// System API/DSM/API/bds_dsm_getDFES_DTC
///This function is used to get DTC values and total number of errors present in DFES entry.
///
///=======
/// Remarks:
///=======
///    + The |GVL_dsm| is given for usage of defines.
///
///----------
/// FFI:
///----------
///This API can be used in trusted partitions only. See Freedom from Interference (FFI) concept for more details.
///
///-----
/// NOTICE:
///-----
///    + On a maximum, 32 different DFES entries are possible. 
///    + Status Mask will take time (max. 10ms) to update in global mask so return status has to be monitored.
///	
///==================================================================		  			===================================================================================================
///Return value    								  									Description
///==================================================================		  			===================================================================================================
///16#0000: BDS_DSM_NO_ERROR_DU16														Update of DTC values and total number of errors present is successful .
///16#0004: BDS_DSM_INVALID_PTR_DU16													Invalid Pointer.
///16#0005: BDS_DSM_MASK_ERROR_DU16													Invalid Mask.
///16#0007: BDS_DSM_INVALID_MAX_ERROR_DU16 											Invalid Max Error.
///16#000B: BDS_DSM_NO_DTC_AVAILABLE_DU16 												Invalid DTC value.
///
///==================================================================		   			===================================================================================================
///
///
///=======
///Code Example:
///=======
///============================================================================
///
///PROGRAM BDS_DSM_getDFES_DTC_TEST
///
///VAR
///
///	mask_s : UINT := BDS_DSM_SET_ACTIVE_ERROR_MASK_DU16;
///
///	startFromBegin_l: BOOL := TRUE;
///
///	maxNum_u16:UINT := 32;
///
///	error_count_u16: UINT;
///
///	dtc_pu16: ARRAY [1..32] OF UINT;
///
///	status_u16: UINT;
///
///END_VAR
///
///dfc_s.id := dfc_ts.DFCid;
///
///(*Get DFES entries*)
///
///status_u16 := bds_dsm_getDFES(mask_s, TRUE, maxNum_u16, ADR(error_count_u16), ADR(dtc_pu16));
///
///if status_u16 = BDS_DSM_NO_ERROR_DU16 THEN
///
///	(*Numbers of Errors have been read successfully*)
///
///END_IF
///
///============================================================================
///
{attribute 'external_name' := 'cmp_rts_bds_dsm_getDFES_DTC'}
FUNCTION bds_dsm_getDFES_DTC : UINT
VAR_INPUT
	///The kind of error status can be specified in detail by means of this mask.
	///
	///Possible values:
	///    + BDS_DSM_SET_ACTIVE_ERROR_MASK_DU16 ( 16#18 ) - Fault is active.
	///    + BDS_DSM_SET_TESTED_ONCE_MASK_DU16 ( 16#08 ) - DFC was tested at least once since start or reset.
	///    + BDS_DSM_SET_TESTED_OK_MASK_DU16 ( 16#20 ) - DFC was at least once ok tested since start or reset.  
	///    + BDS_DSM_SET_FAILED_SINCE_CLEAR_MASK_DU16 ( 16#80 ) - Fault occured at least once since error was deleted from memory.
	mask_s: UINT;
	///
	///    + TRUE: Query is started from the beginning of DFES.
	///    + FALSE: Query is continued with the next index where the last query was finished.
	startFromBegin_l: BOOL;
	///Maximal number of errors/DTCs is returned. The BSW will return at max. 32 values (the max. size of DFES).
	maxNum_u16: UINT;
	///Pointer to a variable where the total number of errors is returned.
	num_pu16: POINTER TO UINT;
	///Pointer variable used to store DTC values.
	dtc_pu16: POINTER TO UINT;
END_VAR

END_FUNCTION

// System API/DSM/API/bds_dsm_getDTC_DFC
///This function returns the DTC of a specified DFC.
///
///=======
/// Remarks:
///=======
///    + The |GVL_dsm| is given for usage of defines.
///	
///----------
/// FFI:
///----------
///This API can be used in trusted partitions only. See Freedom from Interference (FFI) concept for more details.
///
///==================================================================		  			===================================================================================================
///Return value    								  									Description
///==================================================================		  			===================================================================================================
///16#0000: BDS_DSM_NO_ERROR_DU16														Update of DTC of DFC is Successful .
///16#0001: BDS_DSM_DFC_ERROR_DU16														Invalid DFC.
///16#0004: BDS_DSM_INVALID_PTR_DU16													Invalid pointer.
///
///==================================================================		   			===================================================================================================
///
///
///=======
///Code Example:
///=======
///============================================================================
///
///PROGRAM bds_dsm_getDTC_DFC_TEST
///
///VAR
///
///	dfc_s: bds_dsm_dfc_ts;	
///
///	dfc_ts : DFC_bds_NoDebFault1;
///
///	dtc_error_u16 : UINT;
///
///	status_u16: UINT;
///
///END_VAR
///
///dfc_s.id := dfc_ts.DFCid;
///
///(*Read the DTC of DFC*)
///
///dfc_s.id := dfc_ts.DFCid;
///
///status_u16 := bds_dsm_getDTC_DFC(dfc_s,ADR(dtc_error_u16));
///
///if status_u16 = BDS_DSM_NO_ERROR_DU16 THEN
///
///	(*DTC of DFC was read successful*)
///
///END_IF
///
///============================================================================
///
{attribute 'external_name' := 'cmp_rts_bds_dsm_getDTC_DFC'}
FUNCTION bds_dsm_getDTC_DFC : UINT
VAR_INPUT
	///DFC name (identifier) : It is configured using easyConfig tool.
	dfc_s: bds_dsm_dfc_ts;
	///Pointer to a variable where the DTC is returned.
	dtc_pu16: POINTER TO UINT;
END_VAR

END_FUNCTION

// System API/DSM/API/bds_dsm_getDTC_DFCJ1939
///This function is used to read the J1939 specific DTC data (SPN, FMI, Lamp states) for a given DFC.
///
///=======
/// Remarks:
///=======
///    + The |GVL_dsm| is given for usage of defines.
///	+ Suspect Parameter Number (SPN), Failure Mode Identifier (FMI) and Lamp States can be configured in easyConfig.
///	
///----------
/// FFI:
///----------
///This API can be used in trusted partitions only. See Freedom from Interference (FFI) concept for more details.
///
///==================================================================		  			===================================================================================================
///Return value    								  									Description
///==================================================================		  			===================================================================================================
///16#0000: BDS_DSM_NO_ERROR_DU16														Read data is successful.
///16#0001: BDS_DSM_DFC_ERROR_DU16														Wrong DFC.
///16#0004: BDS_DSM_INVALID_PTR_DU16													Invalid Pointer.
///
///==================================================================		   			===================================================================================================
///
///
///=======
///Code Example:
///=======
///============================================================================
///
///PROGRAM bds_dsm_getDTC_DFCJ1939_TEST
///
///VAR
///
///	dfc_s: bds_dsm_dfc_ts;	
///
///	dfc_ts : DFC_bds_NoDebFault1;
///
///	dtcJ1939_s : bds_dsm_dtcj1939_ts;
///
///	status_u16: UINT;
///
///END_VAR
///
///dfc_s.id := dfc_ts.DFCid;
///
///(*Read the DTC of DFC*)
///
///dfc_s.id := dfc_ts.DFCid;
///
///status_u16 := bds_dsm_getDTC_DFCJ1939(dfc_s, ADR(dtcJ1939_s));
///
///if status_u16 = BDS_DSM_NO_ERROR_DU16 THEN
///
///	(*J1939 specific DTC data is read successfull*)
///
///END_IF
///
///============================================================================
///
{attribute 'external_name' := 'cmp_rts_bds_dsm_getDTC_DFCJ1939'}
FUNCTION bds_dsm_getDTC_DFCJ1939 : UINT
VAR_INPUT
	///DFC name (identifier) : It is configured using easyConfig tool.
	dfc_s: bds_dsm_dfc_ts;
	///pointer to a variable where the DTC data is returned.
	dtcJ1939_ps: POINTER TO bds_dsm_dtcj1939_ts;
END_VAR

END_FUNCTION

// System API/DSM/API/bds_dsm_getDTC_J1939
///This function is used to read the J1939 specific DTC data (SPN, FMI, Lamp states) for a given DTC.
///
///=======
/// Remarks:
///=======
///    + The |GVL_dsm| is given for usage of defines.
///	+ Suspect Parameter Number (SPN), Failure Mode Identifier (FMI) and Lamp States can be configured in easyConfig.
///	
///----------
/// FFI:
///----------
///This API can be used in trusted partitions only. See Freedom from Interference (FFI) concept for more details.
///
///----------
/// FFI:
///----------
///This API can be used in trusted partitions only. See Freedom from Interference (FFI) concept for more details.
///
///==================================================================		  			===================================================================================================
///Return value    								  									Description
///==================================================================		  			===================================================================================================
///16#0000: BDS_DSM_NO_ERROR_DU16														Update of J1939 specific data is successful .
///16#0004: BDS_DSM_INVALID_PTR_DU16													Invalid Pointer.
///16#000B: BDS_DSM_NO_DTC_AVAILABLE_DU16												Invalid DTC input.
///
///==================================================================		   			===================================================================================================
///
///
///=======
///Code Example:
///=======
///============================================================================
///
///PROGRAM DSM
///
///VAR
///
///	dfc_s: bds_dsm_dfc_ts;
///
///	dfc_ts : DFC_bds_NoDebFault1;
///
///	dtcJ1939_s: bds_dsm_dtcj1939_ts;
///
///	dtc_u16:UINT := 32772;
///
///	status_u16: UINT;
///
///END_VAR
///
///dfc_s.id := dfc_ts.DFCid;
///
///(*Read the DTC of DFC*)
///
///dfc_s.id := dfc_ts.DFCid;
///
///status_u16 := bds_dsm_getDTC_J1939(dtc_u16, ADR(dtcJ1939_s));
///
///if status_u16 = BDS_DSM_NO_ERROR_DU16 THEN
///
///	(*J1939 specific DTC data is read successfull*)
///
///END_IF
///
///============================================================================
///
///
{attribute 'external_name' := 'cmp_rts_bds_dsm_getDTC_J1939'}
FUNCTION bds_dsm_getDTC_J1939 : UINT
VAR_INPUT
	///DTC value : It is configured using easyConfig tool.
	dtc_u16: UINT;
	///pointer to a variable where the DTC data is returned.
	dtcJ1939_ps: POINTER TO bds_dsm_dtcj1939_ts;
END_VAR

END_FUNCTION

// I/O API/IN legacy/API/bds_in_fi_buffered
///Provides the period array and pulse array of a frequency signal.
///
///=======
/// Remarks:
///=======
///   + In order to receive  the buffered frequency of a signal, it should be configured with easyConfig as a frequency signal. Once configured it is automatically enabled during the start up of the ECU.
///   + For information about the signal acquisition see Frequency acquisition.
///   + If application uses an invalid channel  as a parameter while calling the function, the values stored in the data structure will be 0 // replacement
///   + The following signal information is available: 
///	   + Pointer to the starting address of the Period array (Max size 20).
///	   + Pointer to the starting address of Pulse array (Max size 20).
///   + After the function is called  you get  20  samples of periods and pulses  that could be used within a loop.  
///
///
///----------
/// FFI:
///----------
///This API can be used in trusted partitions only. See Freedom from Interference (FFI) concept for more details.
///
///==================================================================		  			===================================================================================================
///Return value    								  									Description
///==================================================================		  			===================================================================================================
///0																					No error
///1																					Invalid parameter
///2																					Function call was erroneous
///
///==================================================================		   			===================================================================================================
{attribute 'external_name' := 'cmp_rts_bds_in_fi_buffered'}
FUNCTION bds_in_fi_buffered : USINT
VAR_INPUT
	///The signal name that is assigned to the respective pin configured as frequency input. see bds_in_fi_signal_te in bds_rts_ec.xml
	signal_e: UINT;
	///POINTER TO |bds_in_FrqBuffered_ts|
	data_ps: POINTER TO bds_in_FrqBuffered_ts;
END_VAR

END_FUNCTION

// System API/SYS/API/bds_sysPb_getVariant
///This function gets the currently selected post-build selectable variant.
///
///Refer to the page Post-build selectable for more information.
///
///=======
/// Remarks:
///=======
///    + The |GVL_sys| is given for usage of defines.
///    + This Api should be called once in application
///
///----------
/// FFI:
///----------
///This API can be used in trusted partitions.  For untrusted partitions use |bds_sysPb_getVariant_ffi|. See Freedom from Interference (FFI) concept for more details.
///
///==================================================================		  			===================================================================================================
///Return value    								  									Description
///==================================================================		  			===================================================================================================
///|bds_sysPb_retValGetVrnt_ts|															Currently configured variant.
///
///==================================================================		   			===================================================================================================
///
///=======
///Code Example:
///=======
///============================================================================
///
///PROGRAM IniProc
///
///VAR
///	getVaraint_s: bds_sysPb_retValGetVrnt_ts;
///END_VAR
///
///(*getVaraint_s contains the current selected variant*)
///
///getVaraint_s = bds_sysPb_getVariant();
///
///============================================================================
{attribute 'external_name' := 'cmp_rts_bds_sysPb_getVariant'}
FUNCTION bds_sysPb_getVariant : bds_sysPb_retValGetVrnt_ts

END_FUNCTION

// System API/SYS/FFI_API/bds_sysPb_getVariant_ffi
{attribute 'external_name' := 'cmp_rts_bds_sysPb_getVariant_ffi'}
FUNCTION bds_sysPb_getVariant_ffi : bds_sysPb_retValGetVrnt_ts

END_FUNCTION

// System API/SYS/API/bds_sysPb_cfgVariant
///This function is used to select desired variant in the ECU.
///
///Refer to the page Post-build selectable for more information.
///
///=======
/// Remarks:
///=======
///
///The |GVL_sys| is given for usage of defines.
///The selected variant will take effect only after one of the following actions,
///    + A soft reset via bds_sys_resetECU.
///    + Ignition OFF and ON.
///
///----------
/// FFI:
///----------
///This API can be used in trusted partitions only. See Freedom from Interference (FFI) concept for more details.
///
///----------
/// NOTICE:
///----------
///    + The selectable variants will be listed in bds_sysPb_vrnt_te.Import the bds_rts_ec.xml to use the enum.
///    + The configuration related to the particular variant has to be looked-up in easyConfig.
///    + As of now IN module is alone supported for Post-build selectable.
///
///==================================================================		  			===================================================================================================
///Return value    								  									Description
///==================================================================		  			===================================================================================================
///16#0																					No errors, API executed successfully.New variant is updated in RAM successfully.
///16#1																					Invalid variant input.
///16#2																					Variant is already selected
///==================================================================		   			===================================================================================================
///
///=======
///Code Example:
///=======
///============================================================================
///
///PROGRAM IniProc
///
///VAR
///	statusCfgVrnt_s: bds_sysPb_retValCfgVrnt_ts;
///	cfgPbVrnt_u8:usint:=0;
///
///END_VAR
///
///(*Configure a variant. eg bds_sysPb_vrnt03_E*)
///(*Call API once*)
///IF(0 = cfgPbVrnt_u8) THEN
///
///	statusCfgVrnt_s:=bds_sysPb_cfgVariant(bds_sysPb_vrnt_te.bds_sysPb_vrnt03_E);
///
///(*do ignition OFF & ON or do soft reset via bds_sys_resetECU.*)
///cfgPbVrnt_u8:=1;
///
///END_IF
///============================================================================
{attribute 'external_name' := 'cmp_rts_bds_sysPb_cfgVariant'}
FUNCTION bds_sysPb_cfgVariant : bds_sysPb_retValCfgVrnt_ts
VAR_INPUT
	vrntParam_e: USINT;
END_VAR

END_FUNCTION

// I/O API/SENT/API/bds_sent_getFastData
(*The bds_sent_getFastData API function provides the received SENT Fast Data of the selected input signal.

=======
 Remarks:
=======
    + Before accessing the Fast Data frame, check the function call status in the return data structure |bds_sent_rxFastData_ts|.
    + If the function call status is bds_sentCmn_ok_E, then the received Fast Data nibbles from array rxFastData_au8 in the return data structure |bds_sent_rxFastData_ts| can be used. Otherwise the data is set to zero.
    + The function call will return a negative response code if a false parameter is used (e.g., selected signal_e is not defined as SENT input signal or is not configured in Post-Build-Selectable variant).
	+ The positive or negative response codes (e.g., bds_sentCmn_ok_E, bds_sentCmn_notAvl_E and bds_sentCmn_errExt_E) provide in the return data structure |bds_sent_rxFastData_ts| a detailed SENT driver status information chSt_b in bit format.
	+ The number of received Fast Data Nibbles per frame can be configured in easyConfig with the value bds_sent_maxDataNibbles_du8.
	+ The value of the macro define bds_sent_maxDataNibbles_du8 depends on the selected SENT J2716 protocol version. The possible values that can be set in easyConfig are 6 or 8 data nibbles.
	+ The entire SENT channel-specific configuration is to be performed in easyConfig.
	+ Decoding of SENT data is not provided by the API function.

----------
 FFI:
----------
This API can be used in trusted partitions . For untrusted partitions use |bds_sent_getFastData_ffi|. See Freedom from Interference (FFI) concept for more details.
	
==================================================================		  			===================================================================================================
Return value    								  									Description
==================================================================		  			===================================================================================================
|bds_sent_rxFastData_ts|															The return data structure containing the latest received Fast Data sample and the state information.

==================================================================		   			===================================================================================================

=======
Code Example:
=======
============================================================================

PROGRAM appl_10ms_task
VAR

	bds_sent_rxFastData_s : bds_sent_rxFastData_ts;

	idx:USINT;

	appl_sent_rxFastData_au8: ARRAY[1..8] OF USINT;	
	
END_VAR

// Get the single Fast Data frame on selected SENT signal K59

 bds_sent_rxFastData_s = bds_sent_getFastData(bds_sent_signal_te.bds_sent_K59_E);
 
IF(bds_sentCmn_ok_E = bds_sent_rxFastData_s.status_e) THEN
 
    IF(1 = bds_sent_rxFastData_s.chSt_b.newFrmRxd_b1) THEN
   
      // Save the new received Fast Data frame.

      // Received data nibbles saved in low nibble of byte array element (high data nibble set to "0".

		FOR idx := 1 TO 8 BY 1 DO

			appl_sent_rxFastData_au8[idx] := bds_sent_rxFastData_s.rxFastData_au8[idx];

		END_FOR;

    END_IF
  
END_IF

============================================================================

*)
{attribute 'external_name' := 'cmp_rts_bds_sent_getFastData'}
FUNCTION bds_sent_getFastData : bds_sent_rxFastData_ts
VAR_INPUT
	(*The signal name that is assigned to the respective pin configured as SENT channel*)
	signal_e: USINT;
END_VAR

END_FUNCTION

// I/O API/SENT/FFI_API/bds_sent_getFastData_ffi
{attribute 'external_name' := 'cmp_rts_bds_sent_getFastData_ffi'}
FUNCTION bds_sent_getFastData_ffi : bds_sent_rxFastData_ts
VAR_INPUT
	(*The signal name that is assigned to the respective pin configured as SENT channel*)
	signal_e: USINT;
END_VAR

END_FUNCTION

// I/O API/SENT/API/bds_sent_getSlowData
(*The bds_sent_getSlowData API function provides the received SENT Slow Data of the selected input signal.

=======
 Remarks:
=======
    + Before accessing the Slow Data frame, check the function call status in the return data structure |bds_sent_rxSlowData_ts|.
    + If the function call status is bds_sentCmn_ok_E, then the received Slow Data messages from element rxSlowData_u32, msgId_u8 and cfgBit_u8 in the return data structure |bds_sent_rxSlowData_ts| can be used. Otherwise the data is set to zero.
	+ The function call will return a negative response code if a false parameter is used (e.g. selected signal_e is not defined as SENT input signal or is not configured in Post-Build-Selectable variant).
	+ The positive or negative response codes bds_sentCmn_ok_E, bds_sentCmn_notAvl_E and bds_sentCmn_errExt_E support in the return data structure |bds_sent_rxSlowData_ts| a detailed SENT driver status information chSt_b in bit format.
	+ The entire SENT channel-specific configuration is to be performed in easyConfig.
	+ Decoding of SENT data is not provided by the API function.

----------
 FFI:
----------
This API can be used in trusted partitions . For untrusted partitions use |bds_sent_getSlowData_ffi|. See Freedom from Interference (FFI) concept for more details.
	
==================================================================		  			===================================================================================================
Return value    								  									Description
==================================================================		  			===================================================================================================
|bds_sent_rxSlowData_ts|															The return data structure containing the latest received Slow Data sample and the state information

==================================================================		   			===================================================================================================

=======
Code Example:
=======
============================================================================

PROGRAM appl_10ms_task
VAR

	bds_sent_rxSlowData_s : bds_sent_rxSlowData_ts;

	rxSlowData_u32:UDINT;

	SlowData_msgId_u8: USINT;	
	
	SlowData_cfgBit_u8: USINT;
	
END_VAR

// Get the single Slow Data frame on selected SENT signal K59

  bds_sent_rxSlowData_s = bds_sent_getSlowData(bds_sent_signal_te.bds_sent_K59_E);
 
IF(bds_sentCmn_ok_E = bds_sent_rxSlowData_s.status_e) THEN
	
	//Get SENT status information if new Slow Data frame received
 
    IF(1 = bds_sent_rxSlowData_s.chSt_b.newSlowFrmRxd_b1) THEN
   
      // Save the new received Slow Data frame

		rxSlowData_u32 := bds_sent_rxSlowData_s.rxSlowData_u32;

		SlowData_msgId_u8 := bds_sent_rxSlowData_s.msgId_u8;
		
		SlowData_cfgBit_u8 := bds_sent_rxSlowData_s.cfgBit_u8;

	  ELSE

		//error handling for no new Slow Data frame received

    END_IF
  
END_IF

============================================================================

*)
{attribute 'external_name' := 'cmp_rts_bds_sent_getSlowData'}
FUNCTION bds_sent_getSlowData : bds_sent_rxSlowData_ts
VAR_INPUT
	(*The signal name that is assigned to the respective pin configured as SENT channel*)
	signal_e: USINT;
END_VAR

END_FUNCTION

// I/O API/SENT/FFI_API/bds_sent_getSlowData_ffi
{attribute 'external_name' := 'cmp_rts_bds_sent_getSlowData_ffi'}
FUNCTION bds_sent_getSlowData_ffi : bds_sent_rxSlowData_ts
VAR_INPUT
	(*The signal name that is assigned to the respective pin configured as SENT channel*)
	signal_e: USINT;
END_VAR

END_FUNCTION

// I/O API/SENT/API/bds_sent_getFastDataBufd
(*The bds_sent_getFastDataBufd API function provides the latest Buffered Fast Data frame samples from a specified SENT channel.

=======
 Remarks:
=======
    + Before accessing the Buffered Fast Data frame samples, check the function call status in the return data structure |bds_sent_getFastDataBufd_ts|.
    + The number of Buffered Fast Data frame samples can be configured in easyConfig with the value bds_sent_rxFastDataBufSize_du8 from 0 up to maximum 20 number of samples.
    + If the function call status is bds_sentCmn_ok_E, then the received Buffered Fast Data frame samples from array fastDataBufd_as in the return data structure |bds_sent_fastDataMsg_ts| can be used.
	+ The return data structure |bds_sent_fastDataMsg_ts| includes the data array for the Fast Data frame nibbles in the array rxFastData_au8. Otherwise the data is set to zero.
	+ The sequence of the stored Buffered Fast Data frame samples are ordered according LIFO (Last-In-First-Out).
	+ The function call will return a negative response code if a false parameter is used (e.g., selected signal_e is not defined as SENT input signal, is not configured in the Post-Build-Selectable variant or the pointer to the Fast Data buffer fastDataBuf_cps is NULL).
	+ The positive or negative response codes (e.g., bds_sentCmn_ok_E, bds_sentCmn_notAvl_E and bds_sentCmn_errExt_E) provide in the return data structure |bds_sent_getFastDataBufd_ts| a detailed SENT driver status information chSt_b in bit format.
	+ The positive response code bds_sentCmn_ok_E support in the return data structure bds_sent_getFastDataBufd_ts the number of received Buffered Fast Data frames samples cntNewSample_u8 since last function call.
	+ The number of received Fast Data Nibbles per frame can be configured in easyConfig with the value bds_sent_maxDataNibbles_du8.
	+ The value of the macro define bds_sent_maxDataNibbles_du8 depends on the selected SENT J2716 protocol version. The possible values that can be set in easyConfig are 6 or 8 data nibbles.
	+ The entire SENT channel-specific configuration is to be performed in easyConfig.
	+ Decoding of SENT data is not provided by the API function.

----------
 FFI:
----------
This API can be used in trusted partitions . For untrusted partitions use |bds_sent_getFastDataBufd_ffi|. See Freedom from Interference (FFI) concept for more details.
	
==================================================================		  			===================================================================================================
Return value    								  									Description
==================================================================		  			===================================================================================================
|bds_sent_getFastDataBufd_ts|														The return data structure containing the received Fast Data Buffered samples and the state information.

==================================================================		   			===================================================================================================

=======
Code Example:
=======
============================================================================

PROGRAM appl_10ms_task
VAR

	bds_sent_getFastDataBufd_s : bds_sent_getFastDataBufd_ts;

	bds_sent_fastDataBufd_s:bds_sent_fastDataBuf_ts;
	
END_VAR

//Get the Fast Data Buffered frame samples on selected SENT signal K59

bds_sent_getFastDataBufd_s = bds_sent_getFastDataBufd(bds_sent_signal_te.bds_sent_K59_E, ADR(bds_sent_fastDataBufd_s));

============================================================================

*)
{attribute 'external_name' := 'cmp_rts_bds_sent_getFastDataBufd'}
FUNCTION bds_sent_getFastDataBufd : bds_sent_getFastDataBufd_ts
VAR_INPUT
	(*The signal name that is assigned to the respective pin configured as SENT channel*)
	signal_e: USINT;
	(*Pointer to the Fast Data buffered where the data of a particular SENT channel stored*)
	fastDataBuf_cps: POINTER TO bds_sent_fastDataBuf_ts;
END_VAR

END_FUNCTION

// I/O API/SENT/FFI_API/bds_sent_getFastDataBufd_ffi
{attribute 'external_name' := 'cmp_rts_bds_sent_getFastDataBufd_ffi'}
FUNCTION bds_sent_getFastDataBufd_ffi : bds_sent_getFastDataBufd_ts
VAR_INPUT
	(*The signal name that is assigned to the respective pin configured as SENT channel*)
	signal_e: USINT;
	(*Pointer to the Fast Data buffered where the data of a particular SENT channel stored*)
	fastDataBuf_cps: POINTER TO bds_sent_fastDataBuf_ts;
END_VAR

END_FUNCTION

// I/O API/SENT/API/bds_sent_getSlowDataBufd
(*The bds_sent_getSlowDataBufd API function provides the latest Buffered Slow Data frame samples from a specified SENT channel.

=======
 Remarks:
=======
    + Before accessing the Buffered Slow Data frame samples, check the function call status in the return data structure |bds_sent_getSlowDataBufd_ts|.
    + The number of Buffered Slow Data frame samples can be configured in easyConfig with the value bds_sent_rxSlowDataBufSize_du8 from 0 up to maximum 20 number of samples.
    + If the function call status is bds_sentCmn_ok_E, then the received Buffered Slow Data frame samples from array slowDataBufd_as in the return data structure |bds_sent_slowDataMsg_ts| can be used.
	+ The return data structure |bds_sent_slowDataMsg_ts| include the data for the slow Data frame in the element rxSlowData_u32, msgId_u8 and cfgBit_u8. Otherwise the data is set to zero.
	+ The sequence of the stored Buffered Slow Data frame samples are ordered according LIFO (Last-In-First-Out).
	+ The function call will return a negative response code if a false parameter is used (e.g. selected signal_e is not defined as SENT input signal, is not configured in the Post-Build-Selectable variant or the pointer to the Slow Data buffer slowDataBuf_cps is NULL).	+ The function call will return a negative response code if a false parameter is used (e.g., selected signal_e is not defined as SENT input signal, is not configured in the Post-Build-Selectable variant or the pointer to the Fast Data buffer fastDataBuf_cps is NULL).
	+ The positive or negative response codes bds_sentCmn_ok_E, bds_sentCmn_notAvl_E and bds_sentCmn_errExt_E support in the return data structure |bds_sent_getSlowDataBufd_ts| a detailed SENT driver status information chSt_b in bit format.
	+ The positive response code bds_sentCmn_ok_E support in the return data structure |bds_sent_getSlowDataBufd_ts| the number of received Buffered Slow Data frames samples cntNewSample_u8 since last function call.
	+ The entire SENT channel-specific configuration is to be performed in easyConfig.
	+ Decoding of SENT data is not provided by the API function.

----------
 FFI:
----------
This API can be used in trusted partitions . For untrusted partitions use |bds_sent_getSlowDataBufd_ffi|. See Freedom from Interference (FFI) concept for more details.
	
==================================================================		  			===================================================================================================
Return value    								  									Description
==================================================================		  			===================================================================================================
|bds_sent_getSlowDataBufd_ts|														The return data structure containing the received Slow Data Buffered samples and the state information

==================================================================		   			===================================================================================================

=======
Code Example:
=======
============================================================================

PROGRAM appl_10ms_task
VAR

	bds_sent_getSlowDataBufd_s : bds_sent_getSlowDataBufd_ts;

	bds_sent_slowDataBufd_s:bds_sent_slowDataBuf_ts;
	
	appl_sent_cntNewSample_u8: USINT;
	
	cntSavedSamples_u8: USINT;
	
	appl_sent_slowDataBufSamples_s: bds_sent_slowDataBuf_ts;
	
END_VAR

//Get the Slow Data Buffered frame samples on selected SENT signal K59

bds_sent_getSlowDataBufd_s = bds_sent_getSlowDataBufd(bds_sent_signal_te.bds_sent_K59_E, ADR(bds_sent_slowDataBufd_s));

//Check the function call return status

IF(bds_sentCmn_ok_E = bds_sent_getSlowDataBufd_s.status_e) THEN
	
	//check if new Slow Data Buffered frame samples received
	
	appl_sent_cntNewSample_u8 = bds_sent_getSlowDataBufd_s.cntNewSample_u8
 
    IF(0 <> appl_sent_cntNewSample_u8) THEN
   
		FOR cntSavedSamples_u8 := 0 TO appl_sent_cntNewSample_u8 BY 1 DO
			
			//Save the new received Slow Data frame
			
			appl_sent_slowDataBufSamples_s.slowDataBufd_as[cntSavedSamples_u8].rxSlowData_u32 := bds_sent_slowDataBufd_s.slowDataBufd_as[cntSavedSamples_u8].rxSlowData_u32;

			appl_sent_slowDataBufSamples_s.slowDataBufd_as[cntSavedSamples_u8].msgId_u8 := bds_sent_slowDataBufd_s.slowDataBufd_as[cntSavedSamples_u8].msgId_u8;
 
			appl_sent_slowDataBufSamples_s.slowDataBufd_as[cntSavedSamples_u8].cfgBit_u8 := bds_sent_slowDataBufd_s.slowDataBufd_as[cntSavedSamples_u8].cfgBit_u8;

		END_FOR;

	  ELSE

		//error handling for no new Slow Data Buffered frame samples received 

    END_IF
  
END_IF

============================================================================

 *)
{attribute 'external_name' := 'cmp_rts_bds_sent_getSlowDataBufd'}
FUNCTION bds_sent_getSlowDataBufd : bds_sent_getSlowDataBufd_ts
VAR_INPUT
	(*The signal name that is assigned to the respective pin configured as SENT channel*)
	signal_e: USINT;
	(*Pointer to the Slow Data buffered where the data of a particular SENT channel stored*)
	slowDataBuf_cps: POINTER TO bds_sent_slowDataBuf_ts;
END_VAR

END_FUNCTION

// I/O API/SENT/FFI_API/bds_sent_getSlowDataBufd_ffi
{attribute 'external_name' := 'cmp_rts_bds_sent_getSlowDataBufd_ffi'}
FUNCTION bds_sent_getSlowDataBufd_ffi : bds_sent_getSlowDataBufd_ts
VAR_INPUT
	(*The signal name that is assigned to the respective pin configured as SENT channel*)
	signal_e: USINT;
	(*Pointer to the Slow Data buffered where the data of a particular SENT channel stored*)
	slowDataBuf_cps: POINTER TO bds_sent_slowDataBuf_ts;
END_VAR

END_FUNCTION

// I/O API/IN/API/bds_inI_cfgPull
(*The bds_inI_cfgPull provides the option to set the pull type and pull current strength of current inputs.

=======
 Remarks:
=======
	+ The maximum pull current threshold for each input device is 40 mA. If the threshold is exceeded, the API will return bds_inCmn_outOfRng_E.
	+ When shunt resistance is active, switching of pull status is not possible.
	+ Before calling this API, make sure shunt resistance is switched OFF using API |bds_inI_ctrlShunt|.
	+ This API is only applicable for the device inputs refer RC 27-18/40 or RC 18-12/40 Inputs

----------
 FFI:
----------
This API can be used in trusted partitions.For untrusted partitions use |bds_inI_cfgPull_ffi|. See Freedom from Interference (FFI) concept for more details.
	
==================================================================		  			===================================================================================================
Return value    								  									Description
==================================================================		  			===================================================================================================
|bds_inI_cfgPull_ts|																The return structure containing the state information (status_e)

==================================================================		   			===================================================================================================


==================================================================		  			===================================================================================================
Possible status_e values for this function   								  		Description
==================================================================		  			===================================================================================================
bds_inCmn_ok_E																		Call successful and signal can be used
bds_inCmn_invldPrm_E																	+ signal_e is not configured as current input
																						+ pullType or iPull parameter invalid
																						+ Internal device id or channel id invalid
																						+ pullType and iPull combination invalid
bds_inCmn_errInt_E																	Not available due to an internal error
bds_inCmn_errPrecon_E																No valide iPull current selection found. Shunt is not deactivated.
bds_inCmn_invldCfg_E																Requested signal out of range or not configured for active PBS configuration.No default configuration found for iPull current. No stored iPull current found if bds_inCmn_iPull_noChg_E was selected
bds_inCmn_outOfRng_E																The sum current for the device of the signal exceeds max current allowed

==================================================================		   			===================================================================================================

=======
Code Example:
=======
============================================================================

PROGRAM appl_10ms_task
VAR

	pullParam_s : bds_inCmn_pullParam_ts;
	
	cfgPullRtn_s: bds_inI_cfgPull_ts;

END_VAR

// Set the pull type and pull current strength for input A37

cfgPullRtn_s :=  bds_inI_cfgPull(bds_inI_signal_te.bds_inI_A37_E, pullParam_s);

============================================================================

*)
{attribute 'external_name' := 'cmp_rts_bds_inI_cfgPull'}
FUNCTION bds_inI_cfgPull : bds_inI_cfgPull_ts
VAR_INPUT
	(*The signal name that is assigned to the respective pin configured as current input*)
	signal_e: USINT;
	(*Configuration parameters pull type and current strength for current input*)
	pullParam_s: bds_inCmn_pullParam_ts;
END_VAR

END_FUNCTION

// I/O API/IN/API/bds_inI_ctrlShunt
(*The bds_inI_ctrlShunt API function controls the shunt resistor for the input current signal.

=======
 Remarks:
=======
    + Configuration in easyConfig:The inputs supports the reading of analog current if the shunt is activated using easyConfig.
    + Configuration in run time:The shunt resistor of the input must be enabled to measure the analog current.

----------
 FFI:
----------
This API can be used in trusted partitions . For untrusted partitions use |bds_inI_ctrlShunt_ffi|. See Freedom from Interference (FFI) concept for more details.
	
----------
 Info:
----------
    + If the shunt resistor is switched off in run time then voltage measurement is possible for e.g. diagnostic.
	
==================================================================		  			===================================================================================================
Return value    								  									Description
==================================================================		  			===================================================================================================
|bds_inI_shunt_ts|																	The return structure containing the result of control the shunt resistor

==================================================================		   			===================================================================================================

=======
Code Example:
=======
============================================================================

PROGRAM appl_10ms_task
VAR

	bds_inI_ctrlShunt_s : bds_inI_shunt_ts;
	
	bds_inI_getState_s: bds_inI_measmt_ts;

END_VAR

// Control the shunt resistor for the current input signal K30 and switch to OFF

bds_inI_ctrlShunt_s :=  bds_inI_ctrlShunt(bds_inI_Signal_te.bds_inI_K30_E, FALSE);
 
//Get the current information of input signal K30

bds_inI_getState_s = bds_inI_get(bds_inI_Signal_te.bds_inI_K30_E);

============================================================================

*)
{attribute 'external_name' := 'cmp_rts_bds_inI_ctrlShunt'}
FUNCTION bds_inI_ctrlShunt : bds_inI_shunt_ts
VAR_INPUT
	(*The signal name that is assigned to the respective pin configured as current input*)
	signal_e: USINT;
	(*To control the current measurement and the shunt resistor:
    + FALSE: Disable the current measurement and switch OFF the shunt resistor
    + TRUE: Enable the current measurement and switch ON the shunt resistor*)
	cntrl_l: BOOL;
END_VAR

END_FUNCTION

// I/O API/IN/FFI_API/bds_inI_ctrlShunt_ffi
{attribute 'external_name' := 'cmp_rts_bds_inI_ctrlShunt_ffi'}
FUNCTION bds_inI_ctrlShunt_ffi : bds_inI_shunt_ts
VAR_INPUT
	(*The signal name that is assigned to the respective pin configured as current input*)
	signal_e: USINT;
	(*To control the current measurement and the shunt resistor:
    + FALSE: Disable the current measurement and switch OFF the shunt resistor
    + TRUE: Enable the current measurement and switch ON the shunt resistor*)
	cntrl_l: BOOL;
END_VAR

END_FUNCTION

// I/O API/IN/API/bds_inI_get
(*The bds_inI_get API function provides the measurement of the analog current of the input.

=======
 Remarks:
=======
    + Configuration in easyConfig: The inputs supports the reading of analog current if the shunt is activated using easyConfig.
    + Configuration in run time: The |bds_inI_ctrlShunt| API function controls the shunt resistor for the input current signal.
    + The possible measurement range is from 0mA to 24mA.
    + The shunt is protected if the current exceeds 24mA (overcurrent protection), then the shunt is deactivated for a recovery time of 2s. Afterward it is automatically activated again. 

----------
 FFI:
----------
This API can be used in both trusted and untrusted partitions. See Freedom from Interference (FFI) concept for more details.
	
==================================================================		  			===================================================================================================
Return value    								  									Description
==================================================================		  			===================================================================================================
|bds_inI_measmt_ts|																	The return structure containing the current information

==================================================================		   			===================================================================================================

=======
Code Example:
=======
============================================================================

PROGRAM appl_10ms_task
VAR

	bds_inI_getState_s : bds_inI_measmt_ts;

END_VAR

// Get the current information of input signal K30

bds_inI_getState_s := bds_inI_get(bds_inI_Signal_te.bds_inI_K30_E);

============================================================================

*)
{attribute 'external_name' := 'cmp_rts_bds_inI_get'}
FUNCTION bds_inI_get : bds_inI_measmt_ts
VAR_INPUT
	(*The signal name that is assigned to the respective pin configured as current input*)
	signal_e: USINT;
END_VAR

END_FUNCTION

// I/O API/IN/FFI_API/bds_inI_cfgPull_ffi
{attribute 'external_name' := 'cmp_rts_bds_inI_cfgPull_ffi'}
FUNCTION bds_inI_cfgPull_ffi : bds_inI_cfgPull_ts
VAR_INPUT
	(*The signal name that is assigned to the respective pin configured as current input*)
	signal_e: USINT;
	(*Configuration parameters pull type and current strength for current input*)
	pullParam_s: bds_inCmn_pullParam_ts;
END_VAR

END_FUNCTION

// I/O API/IN/API/bds_inDig_get
(*The bds_inDig_get API function provides the measurement of the digital state of the input.

=======
 Remarks:
=======
    + A configuration function is not necessary, because there are no thresholds values to configure.

----------
 FFI:
----------
This API can be used in both trusted and untrusted partition. See Freedom from Interference (FFI) concept for more details.

	
==================================================================		  			===================================================================================================
Return value    								  									Description
==================================================================		  			===================================================================================================
|bds_inDig_measmt_ts|																The return structure containing the digital state information.

==================================================================		   			===================================================================================================

=======
Code Example:
=======
============================================================================

PROGRAM appl_10ms_task
VAR

	bds_inDig_getState_s : bds_inDig_measmt_ts;

	appl_statusDigitalHigh_l:BOOL;

END_VAR

// Get the digital state of input signal K39

bds_inDig_getState_s := bds_inDig_get(bds_inDig_signal_te.bds_inDig_K39_E);

IF (bds_inCmn_ok_E = bds_inDig_getState_s.status_e) THEN

	//save the actual current into local variable

	appl_statusDigitalHigh_l := bds_inDig_getState_s.stHigh_l;

END_IF

============================================================================

*)
{attribute 'external_name' := 'cmp_rts_bds_inDig_get'}
FUNCTION bds_inDig_get : bds_inDig_measmt_ts
VAR_INPUT
	(*The signal name that is assigned to the respective pin configured as digital input*)
	signal_e: USINT;
END_VAR

END_FUNCTION

// I/O API/IN/API/bds_inDig_cfgPull
(*The bds_inDig_cfgPull provides the option to set the pull type and pull current strength of the digital inputs.

=======
 Remarks:
=======
    + The maximum pull current threshold for each input device is 40 mA. If the threshold is exceeded, the API will return bds_inCmn_outOfRng_E.
	+ This API is only applicable for the device inputs refer RC 27-18/40 or RC 18-12/40 Inputs

----------
 FFI:
----------
This API can be used in trusted partitions.  For untrusted partitions use |bds_inDig_cfgPull_ffi|. See Freedom from Interference (FFI) concept for more details.

==================================================================		  			===================================================================================================
Return value    								  									Description
==================================================================		  			===================================================================================================
|bds_inDig_cfgPull_ts|																The return structure containing the state information (status_e)

==================================================================		   			===================================================================================================


==================================================================		  			===================================================================================================
Possible status_e values for this function   								  		Description
==================================================================		  			===================================================================================================
bds_inCmn_ok_E																		Call successful and signal can be used
bds_inCmn_invldPrm_E																	+ signal_e is not configured as digital input
																						+ pullType or iPull parameter invalid
																						+ Internal device id or channel id invalid
																						+ pullType and iPull combination invalid
bds_inCmn_errInt_E																	Not available due to an internal error
bds_inCmn_errPrecon_E																No valide iPull current selection found
bds_inCmn_invldCfg_E																Requested signal out of range or not configured for active PBS configuration.No default configuration found for iPull current. No stored iPull current found if bds_inCmn_iPull_noChg_E was selected
bds_inCmn_outOfRng_E																The sum current for the device of the signal exceeds max current allowed

==================================================================		   			===================================================================================================

=======
Code Example:
=======
============================================================================

PROGRAM appl_10ms_task
VAR

	pullParam_s : bds_inCmn_pullParam_ts;
	
	cfgPullRtn_s: bds_inDig_cfgPull_ts;

END_VAR

// Set the pull type and pull current strength for input K39

cfgPullRtn_s :=  bds_inDig_cfgPull(bds_inDig_signal_te.bds_inDig_K39_E, pullParam_s);

============================================================================

*)
{attribute 'external_name' := 'cmp_rts_bds_inDig_cfgPull'}
FUNCTION bds_inDig_cfgPull : bds_inDig_cfgPull_ts
VAR_INPUT
	(*The signal name that is assigned to the respective pin configured as digital input*)
	signal_e: USINT;
	(*Configuration parameters pull type and current strength for digital input*)
	pullParam_s: bds_inCmn_pullParam_ts;
END_VAR

END_FUNCTION

// I/O API/IN/FFI_API/bds_inDig_cfgPull_ffi
{attribute 'external_name' := 'cmp_rts_bds_inDig_cfgPull_ffi'}
FUNCTION bds_inDig_cfgPull_ffi : bds_inDig_cfgPull_ts
VAR_INPUT
	(*The signal name that is assigned to the respective pin configured as digital input*)
	signal_e: USINT;
	(*Configuration parameters pull type and current strength for digital input*)
	pullParam_s: bds_inCmn_pullParam_ts;
END_VAR

END_FUNCTION

// I/O API/IN/API/bds_inPwm_getTi
(*The bds_inPwm_getTi API function measures the properties of the input PWM signal.

=======
 Remarks:
=======
    + In order to receive the timings of a signal, it shall be configured with easyConfig as a frequency signal.
    + The measurement range of the period time [ns] is defined from 1000000000ns to 50000ns.
    + A call of a configuration function is not required.

----------
 FFI:
----------
This API can be used in trusted partitions . For untrusted partitions use |bds_inPwm_getTi_ffi|. See Freedom from Interference (FFI) concept for more details.
	
==================================================================		  			===================================================================================================
Return value    								  									Description
==================================================================		  			===================================================================================================
|bds_inPwm_tiMeasmt_ts|																The return structure containing the PWM time and state information.

==================================================================		   			===================================================================================================

=======
Code Example:
=======
============================================================================

PROGRAM appl_10ms_task
VAR

	bds_inPwm_getTiPwm_s : bds_inPwm_tiMeasmt_ts;
	
	appl_actualPeriodTime_u32: UDINT;
	
	appl_actualOnWithTime_u32: UDINT;
	
	appl_actualCounterPulse_u32: UDINT;
	
	
END_VAR

// Get the pwm time value of input signal K55

bds_inPwm_getTiPwm_s :=  bds_inPwm_getTi(bds_inPwm_signal_te.bds_inPwm_K55_E);
 
IF (bds_inCmn_ok_E = bds_inPwm_getTiPwm_s.status_e) THEN

    //save the actual pwm times and counter into local variable

    appl_actualPeriodTime_u32   := bds_inPwm_getTiPwm_s.tiPerd_ns_u32;

    appl_actualOnWithTime_u32   := bds_inPwm_getTiPwm_s.tiOnWith_ns_u32;

    appl_actualCounterPulse_u32 := bds_inPwm_getTiPwm_s.cntPls_u32;

END_IF

============================================================================

*)
{attribute 'external_name' := 'cmp_rts_bds_inPwm_getTi'}
FUNCTION bds_inPwm_getTi : bds_inPwm_tiMeasmt_ts
VAR_INPUT
	(*The signal name that is assigned to the respective pin configured as PWM input*)
	signal_e: USINT;
END_VAR

END_FUNCTION

// I/O API/IN/FFI_API/bds_inPwm_getTi_ffi
{attribute 'external_name' := 'cmp_rts_bds_inPwm_getTi_ffi'}
FUNCTION bds_inPwm_getTi_ffi : bds_inPwm_tiMeasmt_ts
VAR_INPUT
	(*The signal name that is assigned to the respective pin configured as PWM input*)
	signal_e: USINT;
END_VAR

END_FUNCTION

// I/O API/IN/API/bds_inPwm_getTiBufd
(*The  bds_inPwm_getTiBufd API function provides a buffered measurement of a PWM signal with up to 20 samples of the input. This can be used to perform an application specific filtering of the PWM data.

=======
 Remarks:
=======
    + In order to receive the buffered timings of a signal, it should be configured with easyConfig as a frequency signal
    + The measured period and time on of the input is given in [ns].
    + The measurement range of the period time [ns] is defined from 1000000000ns to 50000ns.
    + A call of a configuration function is not required.

----------
 FFI:
----------
This API can be used in trusted partitions . For untrusted partitions use |bds_inPwm_getTiBufd_ffi|. See Freedom from Interference (FFI) concept for more details.
	
==================================================================		  			===================================================================================================
Return value    								  									Description
==================================================================		  			===================================================================================================
|bds_inPwm_tiBufd_ts|																The return structure containing the PWM time buffered state.

==================================================================		   			===================================================================================================

=======
Code Example:
=======
============================================================================

PROGRAM appl_10ms_task
VAR

	bds_inPwm_getTiBufd_s : bds_inPwm_tiBufdMeasmt_ts;
	
	bds_inPwm_getTiBufdRet_s : bds_inPwm_tiBufd_ts;
	
	
END_VAR

// Get the pwm time value of input signal K55

  bds_inPwm_getTiBufdRet_s = bds_inPwm_getTiBufd(bds_inPwm_signal_te.bds_inPwm_K55_E,ADR(bds_inPwm_getTiBufd_s));

============================================================================

*)
{attribute 'external_name' := 'cmp_rts_bds_inPwm_getTiBufd'}
FUNCTION bds_inPwm_getTiBufd : bds_inPwm_tiBufd_ts
VAR_INPUT
	(*The signal name that is assigned to the respective pin configured as PWM input*)
	signal_e: USINT;
	(*Pointer to the PWM time buffered information*)
	tiBuf_cps: POINTER TO bds_inPwm_tiBufdMeasmt_ts;
END_VAR

END_FUNCTION

// I/O API/IN/FFI_API/bds_inPwm_getTiBufd_ffi
{attribute 'external_name' := 'cmp_rts_bds_inPwm_getTiBufd_ffi'}
FUNCTION bds_inPwm_getTiBufd_ffi : bds_inPwm_tiBufd_ts
VAR_INPUT
	(*The signal name that is assigned to the respective pin configured as PWM input*)
	signal_e: USINT;
	(*Pointer to the PWM time buffered information*)
	tiBuf_cps: POINTER TO bds_inPwm_tiBufdMeasmt_ts;
END_VAR

END_FUNCTION

// I/O API/IN/API/bds_inR_get
(*The bds_inR_get API function provides the measurement of the resistance of the input.

=======
 Remarks:
=======
    + The measured resistance of the input is given in ohms.
    + The measurement of the resistance range is defined between 20 to 400k ohm and no configuration of the measurement range is needed (700k ohm is the value for an open load or a short circuit to battery).
    + For more information regarding the signal acquisition see Analog voltage acquisition.
    + A call of a configuration function is not required.

----------
 FFI:
----------
This API can be used in both trusted and untrusted partitions. See Freedom from Interference (FFI) concept for more details.
	
==================================================================		  			===================================================================================================
Return value    								  									Description
==================================================================		  			===================================================================================================
|bds_inR_measmt_ts|																	The return structure containing the resistance and state information.

==================================================================		   			===================================================================================================

=======
Code Example:
=======
============================================================================

PROGRAM appl_10ms_task
VAR

	bds_inR_getResistance_s : bds_inR_measmt_ts;
	
	appl_actualResistance_u32: UDINT;

END_VAR

// Get the resistance value of input signal K45

bds_inR_getResistance_s := bds_inR_get(bds_inR_signal_te.bds_inR_K45_E);

IF (bds_inCmn_ok_E = bds_inR_getResistance_s.status_e) THEN

	//save the actual resistance into local variable

	appl_actualResistance_u32 := bds_inR_getResistance_s.r_ohm_u32;

END_IF

============================================================================

*)
{attribute 'external_name' := 'cmp_rts_bds_inR_get'}
FUNCTION bds_inR_get : bds_inR_measmt_ts
VAR_INPUT
	(*The signal name that is assigned to the respective pin configured as resistance input*)
	signal_e: USINT;
END_VAR

END_FUNCTION

// I/O API/IN/API/bds_inPwm_getFrq
(*The bds_inPwm_getFrq API function provides measurement of the frequency of the input signal.

=======
 Remarks:
=======
    + In order to receive the frequency of a signal, it should be configured with easyConfig as a frequency signal
    + The measured frequency of the input is given in [dHz].
    + The measurement range of the frequency [dHz] is defined from 10dHz to 200000dHz.
    + A call of a configuration function is not required.

----------
 FFI:
----------
This API can be used in trusted partitions . For untrusted partitions use |bds_inPwm_getFrq_ffi|. See Freedom from Interference (FFI) concept for more details.
	
==================================================================		  			===================================================================================================
Return value    								  									Description
==================================================================		  			===================================================================================================
|bds_inPwm_frqMeasmt_ts|															The return structure containing the PWM frequency and state information.

==================================================================		   			===================================================================================================

=======
Code Example:
=======
============================================================================

PROGRAM appl_10ms_task
VAR

	bds_inPwm_getFrqPwm_s : bds_inPwm_frqMeasmt_ts;
	
	appl_actualFrequency_u32: UDINT;
	
	appl_actualDutyCycle_Permil_u16: UINT;
	
	appl_actualCounterPulse_u32: UDINT;
	
	appl_counterPulse_LastCall_u32: UDINT;
	
	appl_PulsesPer_10ms_u32: UDINT;
	
END_VAR

//save last pulse counter value

appl_counterPulse_LastCall_u32 := bds_inPwm_getFrqPwm_s.cntPls_u32;

// Get the pwm frequency value of input signal K55

bds_inPwm_getFrqPwm_s :=  bds_inPwm_getFrq(bds_inPwm_signal_te.bds_inPwm_K55_E);
 
IF (bds_inCmn_ok_E = bds_inPwm_getFrqPwm_s.status_e) THEN

    //save the actual pwm times and counter into local variable

    appl_actualFrequency_u32        := bds_inPwm_getFrqPwm_s.frq_dHz_u32;;

    appl_actualDutyCycle_Permil_u16 := bds_inPwm_getFrqPwm_s.dutyCyc_perml_u16;;

    appl_actualCounterPulse_u32     := bds_inPwm_getFrqPwm_s.cntPls_u32;

    //calculate pulses per 10ms

    appl_PulsesPer_10ms_u32 := (appl_actualCounterPulse_u32 - appl_counterPulse_LastCall_u32);

END_IF

============================================================================

*)
{attribute 'external_name' := 'cmp_rts_bds_inPwm_getFrq'}
FUNCTION bds_inPwm_getFrq : bds_inPwm_frqMeasmt_ts
VAR_INPUT
	(*The signal name that is assigned to the respective pin configured as PWM input*)
	signal_e: USINT;
END_VAR

END_FUNCTION

// I/O API/IN/FFI_API/bds_inPwm_getFrq_ffi
{attribute 'external_name' := 'cmp_rts_bds_inPwm_getFrq_ffi'}
FUNCTION bds_inPwm_getFrq_ffi : bds_inPwm_frqMeasmt_ts
VAR_INPUT
	(*The signal name that is assigned to the respective pin configured as PWM input*)
	signal_e: USINT;
END_VAR

END_FUNCTION

// I/O API/IN/API/bds_inU_get
(*The bds_inU_get API function provides the measurement of the analog voltage of the input.

=======
 Remarks:
=======
    + Configuration in easyConfig: The voltage range of the inputs depends on the input type and the input configuration in easyConfig. Based on the configuration, the measurement range of the input can be; Refer to chapter Hardware.
    + Configuration in run time: A call of a configuration function is not required before getting the analog voltage with this bds_inU_get API function.
    + The measurement range of the discrete inputs is 0 to 32000mV and 0 to 5000 mV.
    + The measurement range of the routed input (that means one input of a input device can be routed via the device output directly to the micro controller ADC) via the input device is 0 to 5000mV, see also Analog voltage aquisition.

----------
 FFI:
----------
This API can be used in trusted partitions both trusted and untrusted partitions. See Freedom from Interference (FFI) concept for more details.
	
==================================================================		  			===================================================================================================
Return value    								  									Description
==================================================================		  			===================================================================================================
|bds_inU_measmt_ts|																	The return structure containing the voltage and state information.

==================================================================		   			===================================================================================================

=======
Code Example:
=======
============================================================================

PROGRAM appl_10ms_task
VAR

	bds_inU_getVoltage_s : bds_inU_measmt_ts;
	
	appl_actualVoltage_u16: UINT;

END_VAR

// Get the voltage value of input signal K52

bds_inU_getVoltage_s:=bds_inU_get(bds_inU_signal_te.bds_inU_K52_E);

//get the measured voltage on selected input signal

IF (bds_inCmn_ok_E = bds_inU_getVoltage_s.status_e) THEN

	//save the actual voltage into local variable

	appl_actualVoltage_u16 := bds_inU_getVoltage_s.u_mV_u16;

END_IF

============================================================================

*)
{attribute 'external_name' := 'cmp_rts_bds_inU_get'}
FUNCTION bds_inU_get : bds_inU_measmt_ts
VAR_INPUT
	(*The signal name that is assigned to the respective pin configured as voltage input.*)
	signal_e: USINT;
END_VAR

END_FUNCTION

// I/O API/IN/API/bds_inU_cfgPull
(*The bds_inU_cfgPull function provides the option to set the pull type and pull current strength of the voltage input.

=======
 Remarks:
=======
	+ The maximum pull current threshold for each input device is 40 mA. If the threshold is exceeded, the API will return bds_inCmn_outOfRng_E.
	+ If the voltage input is also configured as current input in easyConfig, then switching pull status shall be controlled by using API |bds_inI_cfgPull|.
	+ If the voltage input is also configured as current input in easyConfig and |bds_inU_cfgPull| is called, then the API returns bds_inCmn_errPrecon_E.
	+ Pull-up 5V doesn't function as expected for 20V and 40V measurement range. 
	+ This API is only applicable for the device inputs refer RC 27-18/40 or RC 18-12/40 Inputs.	

----------
 FFI:
----------
This API can be used in trusted partitions . For untrusted partitions use |bds_inU_cfgPull_ffi|. See Freedom from Interference (FFI) concept for more details.
	
==================================================================		  			===================================================================================================
Return value    								  									Description
==================================================================		  			===================================================================================================
|bds_inU_cfgPull_ts|																The return structure containing the state information (status_e).

==================================================================		   			===================================================================================================


==================================================================		  			===================================================================================================
Possible status_e values for this function    								  		Description
==================================================================		  			===================================================================================================
bds_inCmn_ok_E																		Call successful and signal can be used
bds_inCmn_invldPrm_E																	+ signal_e is not configured as voltage input
																						+ pullType or iPull parameter invalid
																						+ Internal device id or channel id invalid
																						+ pullType and iPull combination invalid
bds_inCmn_errInt_E																	Not available due to an internal error
bds_inCmn_errPrecon_E																No valide iPull current selection found. signal_e is also configured as current input.
bds_inCmn_invldCfg_E																Requested signal out of range or not configured for active PBS configuration.No default configuration found for iPull current. No stored iPull current found if bds_inCmn_iPull_noChg_E was selected
bds_inCmn_outOfRng_E																The sum current for the device of the signal exceeds max current allowed

==================================================================		   			===================================================================================================

=======
Code Example:
=======
============================================================================

PROGRAM appl_10ms_task
VAR

	pullParam_s : bds_inCmn_pullParam_ts;
	
	cfgPullRtn_s: bds_inU_cfgPull_ts;

END_VAR

// Set the pull type and pull current strength for input K52

cfgPullRtn_s :=  bds_inU_cfgPull(bds_inU_signal_te.bds_inU_K52_E, pullParam_s);

============================================================================

*)
{attribute 'external_name' := 'cmp_rts_bds_inU_cfgPull'}
FUNCTION bds_inU_cfgPull : bds_inU_cfgPull_ts
VAR_INPUT
	(*The signal name that is assigned to the respective pin configured as voltage input*)
	signal_e: USINT;
	(*Configuration parameters pull type and current strength for voltage input*)
	pullParam_s: bds_inCmn_pullParam_ts;
END_VAR

END_FUNCTION

// I/O API/IN/FFI_API/bds_inU_cfgPull_ffi
{attribute 'external_name' := 'cmp_rts_bds_inU_cfgPull_ffi'}
FUNCTION bds_inU_cfgPull_ffi : bds_inU_cfgPull_ts
VAR_INPUT
	(*The signal name that is assigned to the respective pin configured as voltage input*)
	signal_e: USINT;
	(*Configuration parameters pull type and current strength for voltage input*)
	pullParam_s: bds_inCmn_pullParam_ts;
END_VAR

END_FUNCTION

// Diagnostics API/UDS/API/bds_uds_registerEvalKeyCallback
///This function registers the callback for Evaluation of Key operation. 
///
///=======
/// Remarks:
///=======
///    + This is the mandatory API to be used to compare the given encrypted response key (e.g. from a diagnostic tool) with the corresponding internal stored and encrypted key for a particular customer configured Security Access Levels. If the keys are equal then the access to the particular security level is provided & its respective callback given will be triggered.
///	   + The callback function is common for all the configured security levels.
///    + The |GVL_uds| is given for usage of defines.
///
///=======
/// INFO:
///=======
///    + The callback will be triggered only if,
///	    + The BODAS security manager is not selected for the security levels in the eC tool.
///	    + Whenever a compare key is requested by a diagnostic tool..
///	   + The customer Instance number zero refers to the BODAS-service Instance and one refers to the ASW customer Instance(customer tool).
///	   + The size of the Key can be configured for a particular security level in the eC tool only if the BODAS security manager is not selected.
///	   + Request seed operation must be done prior to key evaluation.
///	   + The user can configure the security levels using the eC tool. Only levels 1-10 can be configured.
///----------
/// FFI:
///----------
///This API can be used in trusted partitions only. See Freedom from Interference (FFI) concept for more details.
///
///==================================================================		  			===================================================================================================
///Return value    								  									Description
///==================================================================		  			===================================================================================================
///0																					No error
///1																					Invalid pointer
///
///==================================================================		   			===================================================================================================
///
///=======
///Code Example:
///=======
///============================================================================
///
///Callback function
///FUNCTION POU
///VAR_INPUT
///
///    diagInst_u8 : POINTER TO BYTE;(*Diagnostic Instance number*)
///	   secLevel_u8:USINT;(*Security Level.*)
///    key_pau8:POINTER TO USINT;(*Pointer to a buffer which must be provided by the application and which must contain the response key from diagnostic tool for comparison.*)
///    keyLen_u32:USINT;(*Size of key configured in eC*)
///END_VAR
///
///VAR
///	    EvalKeyVar:=usint;
///END_VAR
///
/// To be implemented by the application layer
///IF (EvalKeyVar=0)
///
///  THEN bds_uds_setCallbackStatus(0);(*positive response*)
///  
///END_IF
///
///IF (EvalKeyVar=1) 
///
///  THEN  bds_uds_setCallbackStatus(1);(*negative response*)
///  
///END_IF
///IF (EvalKeyVar=2)
///
///  THEN bds_uds_setCallbackStatus(16#B);(*Key is incorrect or not matching with calculated Key.*)
///  
///END_IF
///
///IF (EvalKeyVar=3) 
///
///  THEN  bds_uds_setCallbackStatus(16#10);(*This asynchronous function was not yet completed and must be called again with the same parameter values.*)
///  
///END_IF
///
///(*Registering callback*)
///
///PROGRAM POU_10
///VAR
///
///	flag_1 : usint := 0;
///
///END_VAR
///
///IF ( flag_1=0)
///
///    THEN bds_uds_registerEvalKeyCallback (ADR(POU));
///
///    flag_1 := 1;(*To make api call once in application*)
///
///END_IF
///
///
///============================================================================
{attribute 'external_name' := 'cmp_rts_bds_uds_registerEvalKeyCallback'}
FUNCTION bds_uds_registerEvalKeyCallback : USINT
VAR_INPUT
	///Function pointer with argument as mentioned above
	func_pf: POINTER TO BOOL;
END_VAR

END_FUNCTION

// Diagnostics API/UDS/API/bds_uds_registerGetSeedCallback
///This function registers the callback for Get seed operation. 
///
///=======
/// Remarks:
///=======
///    + This is the mandatory API to be used to request a seed value for a particular customer configured security level.
///	   + The callback function is common for all the configured security levels.
///    + The |GVL_uds| is given for usage of defines.
///
///=======
/// INFO:
///=======
///    + The callback will be triggered only if,
///	    + The BODAS security manager is not selected for the security levels in the eC tool.
///	    + Whenever a seed is requested by a diagnostic tool.
///	   + The customer Instance number zero refers to the BODAS-service Instance and one refers to the ASW customer Instance(customer tool).
///	   + The size of the Seed can be configured for a particular security level in the eC tool only if the BODAS security manager is not selected.
///	   + The user can configure the security levels using the eC tool. Only levels 1-10 can be configured.
///----------
/// FFI:
///----------
///This API can be used in trusted partitions only. See Freedom from Interference (FFI) concept for more details.
///
///==================================================================		  			===================================================================================================
///Return value    								  									Description
///==================================================================		  			===================================================================================================
///0																					No error
///1																					Invalid pointer
///
///==================================================================		   			===================================================================================================
///
///=======
///Code Example:
///=======
///============================================================================
///
///Callback function
///FUNCTION POU
///VAR_INPUT
///
///    diagInst_u8 : POINTER TO BYTE;(*Diagnostic Instance number*)
///	   secLevel_u8:USINT;(*Security Level.*)
///    seed_pau8:POINTER TO USINT;(*Pointer to a buffer which must be provided by the application. Generated seed will be copied to this buffer.*)
///    seedLen_u32:USINT;(*Size [in bytes] of the seed configured in eC.*)
///END_VAR
///
///VAR
///	    getSeedVar:=usint;
///END_VAR
///
/// To be implemented by the application layer
///IF (getSeedVar=0)
///
///  THEN bds_uds_setCallbackStatus(0);(*positive response*)
///  
///END_IF
///
///IF (getSeedVar=1) 
///
///  THEN  bds_uds_setCallbackStatus(1);(*negative response*)
///  
///END_IF
///
///IF (getSeedVar=3) 
///
///  THEN  bds_uds_setCallbackStatus(16#10);(*This asynchronous function was not yet completed and must be called again with the same parameter values.*)
///  
///END_IF
///
///(*Registering callback*)
///
///PROGRAM POU_10
///VAR
///
///	flag_1 : usint := 0;
///
///END_VAR
///
///IF ( flag_1=0)
///
///    THEN bds_uds_registerGetSeedCallback (ADR(POU));
///
///    flag_1 := 1;(*To make api call once in application*)
///
///END_IF
///
///
///============================================================================
{attribute 'external_name' := 'cmp_rts_bds_uds_registerGetSeedCallback'}
FUNCTION bds_uds_registerGetSeedCallback : USINT
VAR_INPUT
	///Function pointer with argument as mentioned above
	func_pf: POINTER TO BOOL;
END_VAR

END_FUNCTION

// System API/SYS/API/bds_sys_applSwName
///This function updates the application software name. By default, the application software name is 'CodesysApplication'.
///
///----------
/// FFI:
///----------
///This API can be used in trusted partitions only.
///	
///==================================================================		  			===================================================================================================
///Return value    								  										Description
///==================================================================		  			===================================================================================================
///|bds_sys_retValApplSwName_ts|														The return structure containing the function call status (status_e). 
///
///==================================================================		   			===================================================================================================
///
///==================================================================		  			===================================================================================================
///Possible status_e values for this function    								  		Description
///==================================================================		  			===================================================================================================
///bds_sys_swnmOk_E																		Function is called without errors.
///bds_sys_errSwnm_E																	String length of ASW name is too long / invalid parameter.
///
///==================================================================		   			===================================================================================================
///
///=======
///Code Example:
///=======
///============================================================================
///
///PROGRAM appl_10ms_task
///
///VAR
///
///	applSwName_au8:STRING(50):='TestApplication';
///
///	retValApplSwName_s : bds_sys_retValApplSwName_ts;
///
///END_VAR
///
///
///(* update the application software name *)
///
/// retValApplSwName_s:=bds_sys_applSwName(ADR(applSwName_au8));
///
///
///============================================================================
{attribute 'external_name' := 'cmp_rts_bds_sys_applSwName'}
FUNCTION bds_sys_applSwName : bds_sys_retValApplSwName_ts
VAR_INPUT
	applSwName_pau8: POINTER TO STRING(50);(*Pointer to a character string with software name. The max string length is 50 characters (chars).*)
END_VAR

END_FUNCTION

// I/O API/OUT/API/bds_outClcU_rstErr
/// The BODAS API-Function resets an existing diagnostic fault error and reactivating of voltage outputs, which are switched off due to an error detection.
///
///=======
///----------
/// FFI:
///----------
/// This API can be used in trusted partitions. For untrusted partitions use bds_outClcU_rstErr_ffi. See Freedom from Interference (FFI) concept for more details.
///
///
///==================================================================		  			===================================================================================================
///Return value    								  									    Description
///==================================================================		  			===================================================================================================
///bds_outClcU_rstErr_ts														        The return structure containing the state information (statusApi_e)
///
///==================================================================		   			===================================================================================================
///
///=======
///Code Example:
///=======
///============================================================================
///
/// PROGRAM appl_10ms_task
/// VAR
///     bds_outClcU_signal_e : bds_outClcU_signal_te;
///     bds_outClcU_retRstErr_s : bds_outClcU_rstErr_ts;
/// END_VAR
/// 
/// bds_outClcU_signal_e := bds_outClcU_signal_te.bds_outClcU_K25_E;
/// 
/// (* call BDS-Function *)
/// bds_outClcU_retRstErr_s := bds_outClcU_rstErr(bds_outClcU_signal_e);
/// 
/// IF bds_outCmn_ok_E = bds_outClcU_retRstErr_s.statusApi_e THEN
///     (* Call successful, signal is valid *)
///     (* reset of an existing diagnostic fault error and reactivating of voltage outputs *)
/// ELSE
///     (* error handling *)
/// END_IF
/// END_PROGRAM
///
///============================================================================
{attribute 'external_name' := 'cmp_rts_bds_outClcU_rstErr'}
FUNCTION bds_outClcU_rstErr : bds_outClcU_rstErr_ts
VAR_INPUT
	///The connector assigned signal name of the output.
	signal_e: USINT;
END_VAR

END_FUNCTION

// I/O API/OUT/API/bds_outDig_set
///The BODAS API-Function set the digital output to particular state.
///
///=======
/// Remarks:
///=======
/// The threshold FOR the over current detection FOR high power digital outputs is 6500[mA].

/// Set the digital output state for all "Highside High power outputs", "Lowside High power outputs" and "Lowside Low power outputs" (available signal refer to RC27-18/40 - Outputs).

///FOR more information see topic Digital outputs.

///
///----------
/// FFI:
///----------
///This API can be used in trusted partitions. For untrusted partitions use bds_outDig_set_ffi. See Freedom from Interference (FFI) concept for more details.
///
///------
/// Info:
///------
///
/// +Macro define "bds_outDig_endNumSigDig_D" in easyConfig generated file "bds_outDig_ec.h" defines the end of the Digital output signals in the digital enumeration type definition "bds_outDig_signal_te".
/// 
/// +Macro define "bds_outDig_strtNumSigPwm_D" in easyConfig generated file "bds_outDig_ec.h" defines the start of the Pwm output signals if used in digital mode ( OFF = 0% and ON = 100% duty cycle).

///
///Attention
 
/// +It is possible to poll the status of the fault. If the error has been healed, then the output can be unlocked by calling this API-Function.

/// +After a hot short circuit and over current the unlock of the high power output is only possible after a reactivation wait time of 2s, refer to bit in status bds_outCmn_statusDiag_tb.
 
///
///==================================================================		  			===================================================================================================
///Return value    								  									    Description
///==================================================================		  			===================================================================================================
///bds_outDig_set_ts															        The return structure containing the state information (statusApi_e)
///
///==================================================================		   			===================================================================================================
///
///=======
///Code Example:
///=======
///============================================================================
///
///Set digital output pin to ON
/// 
/// PROGRAM appl_10ms_task
///
/// VAR
///
///     bds_outDig_signal_e : bds_outDig_signal_te;
///
///     bds_outDig_retSet_s : bds_outDig_set_ts;
///
///     flgEna_l : BOOL;
///
/// END_VAR
/// 
/// bds_outDig_signal_e := bds_outDig_signal_te.bds_outDig_K13_E;
///
/// flgEna_l := TRUE;
/// 
/// (* call BDS-Function *)
///
/// bds_outDig_retSet_s := bds_outDig_set(bds_outDig_signal_e, flgEna_l);
/// 
/// IF bds_outCmn_ok_E = bds_outDig_retSet_s.statusApi_e THEN
///
///     (* Call successful, signal is valid *)
///
///     (* set the digital output to requested state *)
///
/// ELSE
///
///     (* error handling *)
///
/// END_IF
///
/// END_PROGRAM
/// 
/// Set PWM signal used as digital output pin to ON
///
/// PROGRAM appl_10ms_task
///
/// VAR
///
///     bds_outDig_signal_e : bds_outDig_signal_te;
///
///     bds_outDig_retSet_s : bds_outDig_set_ts;
///
///     flgEna_l : UINT;
///
/// END_VAR
/// 
/// bds_outDig_signal_e := bds_outDig_K07_E;
///
/// flgEna_l := 1;
/// 
/// (* call BDS-Function *)
///
/// bds_outDig_retSet_s := bds_outDig_set(bds_outDig_signal_e, flgEna_l);
/// 
/// IF bds_outCmn_ok_E = bds_outDig_retSet_s.statusApi_e THEN
///
///     (* Call successful, signal is valid *)
///
///     (* set the digital output to requested state *)
///
/// ELSE
///
///     (* error handling *)
///
/// END_IF
///
/// END_PROGRAM
///
///============================================================================
{attribute 'external_name' := 'cmp_rts_bds_outDig_set'}
FUNCTION bds_outDig_set : bds_outDig_set_ts
VAR_INPUT
	///The connector assigned signal name of the output.
	signal_e: USINT;
	/// defining the digital state of the selected digital output signal (FALSE = OFF, TRUE = ON)
	flgEna_l: BOOL;
END_VAR

END_FUNCTION

// I/O API/OUT/API/bds_outDig_get
///The BODAS API-function gets the detailed status information of the digital output as well as PWM signals used as digital output.
///
///=======
/// Remarks:
///=======
/// The "current measurement" AND corresponding "current sensing" is just possible FOR the "high power outputs".

/// The threshold for the over current detection is 6500mA and therefore also the measurement range is defined from 0 to 6500mA.

/// The status data holds all relevant information of the digital output, see the example below.

/// Part of the status bit field is also the fault error status of every DFC (e.g. stErrSCB_b1), see topic Digital outputs and Diagnostic Fault Check. 


///
///----------
/// FFI:
///----------
/// This API can be used in both trusted and untrusted partitions. See Freedom from Interference (FFI) concept for more details.
///
///------
///
///==================================================================		  			===================================================================================================
///Return value    								  									    Description
///==================================================================		  			===================================================================================================
///bds_outDig_get_ts														            The return structure containing:
///																							- The digital state ON or OFF of the digital output
///																							- The measured current value of the digital output in [mA]
///																							- Detailed diagnostic information of the digital output
///																							- Function call status information (statusApi_e)

///
///==================================================================		   			===================================================================================================
///
///=======
///Code Example:
///=======
///============================================================================
///
/// PROGRAM appl_10ms_task
///
/// VAR
///
///     bds_outDig_signal_e : bds_outDig_signal_te;
///
///     bds_outDig_retGet_s : bds_outDig_get_ts;
///
///     retVal_stFlgEna_l : BOOL;
///
///     retVal_iAct_mA_u16 : UINT;
///
/// END_VAR
/// 
/// bds_outDig_signal_e := bds_outDig_signal_te.bds_outDig_K13_E;
/// 
/// (* call BDS-Function - Set digital output state *)
///
/// bds_outDig_set(bds_outDig_signal_e, TRUE);
/// 
/// (* call BDS-Function - Get status and diagnostic information *)
///
/// bds_outDig_retGet_s := bds_outDig_get(bds_outDig_signal_e);
/// 
/// IF bds_outCmn_ok_E = bds_outDig_retGet_s.statusApi_e THEN
///
///     (* Call successful, signal is valid *)
///
///     (* check if there is a short cut to battery or to ground? *)
///
///     IF (TRUE = bds_outDig_retGet_s.statusDiag_b.stErrSCB_b1) OR (TRUE = bds_outDig_retGet_s.statusDiag_b.stErrSCG_b1) THEN
///
///         (* SCB or SCG - Set values to zero *)
///
///         retVal_stFlgEna_l := FALSE;
///
///         retVal_iAct_mA_u16 := 0;
///
///     ELSE
///
///         (* get digital state on requested output *)
///
///         retVal_stFlgEna_l := bds_outDig_retGet_s.stFlgEna_l;
///
///         (* get actual measured current on requested output *)
///
///         retVal_iAct_mA_u16 := bds_outDig_retGet_s.iAct_mA_u16;
///
///     END_IF
///
/// ELSE
///
///     (* error handling *)
///
/// END_IF
///
/// END_PROGRAM
///
///============================================================================
{attribute 'external_name' := 'cmp_rts_bds_outDig_get'}
FUNCTION bds_outDig_get : bds_outDig_get_ts
VAR_INPUT
	///The connector assigned signal name of the output.
	signal_e: USINT;
END_VAR

END_FUNCTION

// I/O API/OUT/API/bds_outDig_cfgDiag
/// The BODAS API-function configure the diagnostic features of the selected digital output as well as PWM signals used as digital output.
/// 
/// ·Control the full diagnostic of selected digital output
/// 
/// ·Control the selected digital output and set to unused and disable the diagnosis
/// 
/// ·Control the open load detection of the selected digital output
/// 
/// ·Control the detection of non hot short circuit error of the selected digital output

///
///=======
/// Remarks:
///=======
///
/// +Control the full diagnostic of selected digital output:
///
/// +Test pulses are enabled by default.
///
/// +For some application this test pulses disturb the wanted functionality of the output for example if you want to use it for power supply.
///
/// +The test pulses can be deactivated for High Power Outputs only.
///Attention 
///
///If test pulses are disabled, for an output then the fault detection and healing is limited. Please refer to topic Digital outputs

/// + Control the selected digital output and set to unused and disable the diagnosis:
/// 
/// + Disable an unused output and its diagnosis.
/// 
/// + The output should be disabled during start up.
/// Attention
///If an output is disabled, faults are not longer detected and also the diagnostic control of the output is disabled.

/// +Control the open load detection of high side and low side digital output:
/// 
/// +Open load detection is enabled by default. Hence it can be disabled and enabled for the digital high side or low side output.
///
/// +If open load detection is disabled, Open load will not be detected and healed.
///
/// +For example in some application the open load detection may disturb the required functionality of an output. For example if the high power high side digital output is used as power supply for the low side digital output.
///
/// +Please refer topic Digital outputs for open load detection of digital high side and low side output. 
///
/// +Control the non-hot short circuit detection of high side and low side digital output:
///
/// +Non hot short circuit detection is enabled by default. Hence it can be disabled and enabled for the PWM high side or low side output.
///
/// +If non hot short circuit detection is disabled, Non hot short circuit will not be detected and healed.
///
/// +For high side digital output short circuit to battery is non hot error and for low side digital output short circuit to ground is non hot error.
///
/// +Please refer topic Digital outputs for non hot short circuit detection of digital high side and low side output. 
 
///----------
/// FFI:
///----------
///This API can be used in trusted partitions. For untrusted partitions use bds_outDig_cfgDiag_ffi. See Freedom from Interference (FFI) concept for more details.
///
///------
/// Info:
///------
/// Diagnostic configurations shall be disabled during start up of the application, otherwise faults may be detected on the time of diagnostic configuration. The previously detected faults can be reset with bds_outDig_rstErr.

/// For more information, refer to bds_outDig_get.
 
/// The return structure member "statusDiag_b" holds the information regarding the configuration.

///
///Attention
 
/// +It is possible to poll the status of the fault. If the error has been healed, then the output can be unlocked by calling this API-Function.
///
/// +After a hot short circuit and over current the unlock of the high power output is only possible after a reactivation wait time of 2s, refer to bit in status bds_outCmn_statusDiag_tb.
 
///
///==================================================================		  			===================================================================================================
///Return value    								  									    Description
///==================================================================		  			===================================================================================================
///bds_outDig_cfgDiag_ts														        The return structure containing the state information (statusApi_e)
///
///==================================================================		   			===================================================================================================
///
///=======
///Code Example:
///=======
///============================================================================
///
/// PROGRAM OsIniProc
///
/// VAR
///
///     bds_outDig_signal_e : bds_outDig_signal_te;
///
///     bds_outDig_retCfgDiag_s : bds_outDig_cfgDiag_ts;
///
///     diagParam_s : bds_outCmn_diagParam_ts;
///
/// END_VAR
/// 
/// bds_outDig_signal_e := bds_outDig_signal_te.bds_outDig_K13_E;
/// 
/// (* configure the diagnostic feature of the digital output *)
///
/// diagParam_s.diFullDiag_l := FALSE;
///
/// diagParam_s.diCntlAndDiag_l := TRUE;
///
/// diagParam_s.diOpenLoadDetn_l := FALSE;
///
/// diagParam_s.diNonHotSCDetn_l := FALSE;
/// 
/// (* call BDS-Function - Configure the diagnostic feature for the requested digital output *)
///
/// bds_outDig_retCfgDiag_s := bds_outDig_cfgDiag(bds_outDig_signal_e, diagParam_s);
/// 
/// IF bds_outCmn_ok_E = bds_outDig_retCfgDiag_s.statusApi_e THEN
///
///     (* Call successful, signal is valid *)
///
///     (* Disabled the output and the diagnosis for this requested digital output *)
/// ELSE
///
///     (* error handling *)
///
/// END_IF
///
/// END_PROGRAM
///============================================================================
{attribute 'external_name' := 'cmp_rts_bds_outDig_cfgDiag'}
FUNCTION bds_outDig_cfgDiag : bds_outDig_cfgDiag_ts
VAR_INPUT
	///The connector assigned signal name of the output.
	signal_e: USINT;
	/// defining the digital state of the selected digital output signal (FALSE = OFF, TRUE = ON)
	diagParam_s: bds_outCmn_diagParam_ts;
END_VAR

END_FUNCTION

// I/O API/OUT/API/bds_outDig_rstErr
/// The BODAS API-function reset the diagnostics error and unlocks the digital outputas well as PWM signals used as digital output.
///=======
/// Remarks:
///=======
///  +After a fault the digital output is locked but the set point is still valid. With the error is reset, output is also unlocked.
///  
///  +After a hot short circuit and over current the unlocking of the power output is only possible after a reactivation time of 2s.
///  
///  +It is possible to poll the status of the fault. If the error has been healed, then the output can be reset.
///  
///  +For over current fault: After reset, the output has to be switched on again using the API bds_outDig_set.
///  
///  +For more information see topic Digital outputs.

///----------
/// FFI:
///----------
/// This API can be used in trusted partitions. For untrusted partitions use bds_outDig_rstErr_ffi. See Freedom from Interference (FFI) concept for more details.
///
///
///==================================================================		  			===================================================================================================
///Return value    								  									    Description
///==================================================================		  			===================================================================================================
///bds_outDig_rstErr_ts														            The return structure containing the state information (statusApi_e)
///
///==================================================================		   			===================================================================================================
///
///=======
///Code Example:
///=======
///============================================================================
///
/// PROGRAM appl_10ms_task
///
/// VAR
///
///     bds_outDig_signal_e: bds_outDig_signal_te; 
///
///     bds_outDig_retRstErr_s: bds_outDig_rstErr_ts;
///
/// END_VAR
/// 
/// bds_outDig_signal_e := bds_outDig_signal_te.bds_outDig_K13_E; (* Assigning a specific signal*)
/// 
/// (* Calling a function to reset the diagnostic error and unlock the digital output*)
///
/// bds_outDig_retRstErr_s := bds_outDig_rstErr(bds_outDig_signal_e);
/// 
///   (*Checking the return state of the function call*)
///
/// IF bds_outCmn_ok_E = bds_outDig_retRstErr_s.statusApi_e THEN
///
///       (*Call successful, signal is valid*)
///
///      (*Reset the diagnostics error and unlocks the digital output*)
///
/// ELSE
///
///      (*Handle the error*)
///
/// END_IF;
/// 
/// END_PROGRAM
///
///============================================================================
{attribute 'external_name' := 'cmp_rts_bds_outDig_rstErr'}
FUNCTION bds_outDig_rstErr : bds_outDig_rstErr_ts
VAR_INPUT
	///The connector assigned signal name of the output.
	signal_e: USINT;
END_VAR

END_FUNCTION

// I/O API/OUT/API/bds_outPwm_setDutyCycle
///The BODAS API-function sets the PWM high side or low side output with different range of duty cycles from 0% up to 100%.
///
///=======
/// Remarks:
///=======
/// After a fault the output is locked but the set point is still valid.
/// For more information see topic Proportional outputs.
/// Attention
/// It is possible to poll the status of the fault. If the error has been healed, then the output can be unlocked by calling this API-Function.
/// After a hot short circuit and over current the unlock of the high power output is only possible after a reactivation wait time of 2s, refer to bit in status bds_outCmn_statusDiag_tb.
 
///
///----------
/// FFI:
///----------
/// This API can be used in trusted partitions. For untrusted partitions use bds_outPwm_setDutyCycle_ffi. See Freedom from Interference (FFI) concept for more details.
///
///------
///
///==================================================================		  			===================================================================================================
///Return value    								  									    Description
///==================================================================		  			===================================================================================================
///bds_outPwm_setDutyCycle_ts														            The return structure containing the state information (statusApi_e)
///
///==================================================================		   			===================================================================================================
///
///=======
///Code Example:
///=======
///============================================================================
///
/// PROGRAM appl_10ms_task
///
///VAR
///
///    bds_outPwm_signal_e: bds_outPwm_signal_te;
///	
///    bds_outPwm_retSetDutyCycle_s: bds_outPwm_setDutyCycle_ts;
///	
///    ratDutyCycle_perml_u16: UINT := 500; (* 500 is 50% duty cycle with 0.1% resolution *)
///	
///END_VAR
///
///bds_outPwm_signal_e := bds_outPwm_signal_te.bds_outPwm_K09_E;
///
///(* Call BDS-Function to actuate output with duty-cycle *)
///
///bds_outPwm_retSetDutyCycle_s := bds_outPwm_setDutyCycle(bds_outPwm_signal_e, ratDutyCycle_perml_u16);
///
///(* check return state of BDS-Function call *)
///
///IF bds_outCmn_ok_E = bds_outPwm_retSetDutyCycle_s.statusApi_e THEN
///
///    (* Call successful, signal is valid *)
///	
///    (* Actuated the Pwm output to requested duty-cycle successfully *)
///	
///ELSE
///
///    (* error handling *)
///	
///END_IF
///
/// END_PROGRAM
///============================================================================
{attribute 'external_name' := 'cmp_rts_bds_outPwm_setDutyCycle'}
FUNCTION bds_outPwm_setDutyCycle : bds_outPwm_setDutyCycle_ts
VAR_INPUT
	///The connector assigned signal name of the output.
	signal_e: USINT;
	///The connector assigned signal name of the output.
	ratDutyCycle_perml_u16: UINT;
END_VAR

END_FUNCTION

// I/O API/OUT/API/bds_outPwm_get
///The BODAS API-function gets the detailed status of a PWM high side or low side output.
///
///=======
/// Remarks:
///=======
///The threshold FOR the over current detection is 6500mA AND therefore also the measurement range is defined FROM 0..6500mA.
///
///The status data holds all relevant information of the proportional output, see example below.
///
///Part of the status bit field is also the fault error status of every DFC (e.g. stErrSCB_b1). See  the topic Proportional outputs and Diagnostic Fault Check. 
 
